(*
    This function runs all test suites that have been initialized.
    The test suites are run in parallel (all at once).
*)
FUNCTION RUN

GVL_TcUnit.TcUnitRunner.RunTestSuiteTests();

END_FUNCTION

(* stored: Version 1.1.0.1
   POU RUN: Id {bd49b256-e7ba-4b73-b669-380d1f428417}, SpecialFunc None *)
